// TIA Portal V20 export
VAR_GLOBAL   // PLC tag table "PLC-A3-DI"
   "ENCODER_L+" AT %I0.0 : Bool;   // JEDEN ENCODER DVA KANÁLY NAASTAVENÍ NA HSPEED COUNTER
   "ENCODER_L-" AT %I0.1 : Bool;   // JEDEN ENCODER DVA KANÁLY NAASTAVENÍ NA HSPEED COUNTER
   ENCODER AT %I0.2 : Bool;
   "ENCODER(1)" AT %I0.3 : Bool;
   "ENCODER(2)" AT %I0.4 : Bool;
   RESERVE_DI AT %I0.5 : Bool;   // s1 najezd
   RESERVE_DI_1 AT %I0.6 : Bool;   // s2 foceni
   RESERVE_DI_2 AT %I0.7 : Bool;   // s3 konec budky
   RESERVE_DI_3 AT %I1.0 : Bool;   // s4 vyrazovač
   RESERVE_DI_4 AT %I1.1 : Bool;   // s5 valec pozice home
   RESERVE_DI_5 AT %I1.2 : Bool;
   RESERVE_DI_6 AT %I1.3 : Bool;
   RESERVE_DI_7 AT %I1.4 : Bool;
   RESERVE_DI_8 AT %I1.5 : Bool;
END_VAR
